{attribute 'qualified_only'}
{attribute 'strict'}
{attribute 'to_string'}
TYPE E_HomeIndexState :
(
    Idle := 0,
    Homing,
    WaitHomed,
    HomingUnlatch,
    HomingPulsed,
    WaitHomeDone,
    CenterMove,
    WaitCenterDone,
    SetPosition,
    HomingDone,
    Done,
    Error
)UINT;
END_TYPE

(* stored: Version 1.1.0.1
   DUT E_HomeIndexState: Id {736988bd-d907-4bb5-b974-c2963365e1d6} *)
